Fanuc KAREL source: KT00865.KL

PROGRAM KT00865
%NOLOCKGROUP
VAR
  B1: BOOLEAN
  B2: BOOLEAN
  OUT: REAL
BEGIN
  B1 = TRUE
  B2 = FALSE
  B1 = TRUE
  B2 = FALSE
  OUT = ROUND(B1)
END KT00865
